(* IEC 61131-3 sources: plc-process-lib/src/POUs/Time/FB_FakeTime, 4 files *)

(* ---- FB_FakeTime.decl.st ---- *)
// Назначение: подменяемый источник времени для тестов: время меняется только вызовами
//             SetNow, Advance, AdvanceL, поэтому тесты таймингов детерминированы и не ждут
//             реального времени. Лежит в библиотеке (не в tests/): им пользуются тесты
//             проектов-потребителей. Старт — LTIME#1H, а не 0: ловит код, который считает
//             «0 = не инициализировано».
// Автор:      kr0nsch
// Версия:     0.1.0
// Документ:   docs/fb/FB_FakeTime.md
FUNCTION_BLOCK FB_FakeTime IMPLEMENTS I_TimeSource
VAR
    ltNow : LTIME := LTIME#1H;   // текущее подменное время
END_VAR

(* ---- Advance.method.decl.st ---- *)
// Продвинуть время на шаг TIME (мс)
METHOD PUBLIC Advance
VAR_INPUT
    tStep : TIME;   // шаг
END_VAR

(* ---- AdvanceL.method.decl.st ---- *)
// Продвинуть время на шаг LTIME: шаги меньше 1 мс и больше 49 сут
METHOD PUBLIC AdvanceL
VAR_INPUT
    ltStep : LTIME;   // шаг
END_VAR

(* ---- SetNow.method.decl.st ---- *)
// Установить время. Можно и назад: ФБ библиотеки обязаны это переживать
METHOD PUBLIC SetNow
VAR_INPUT
    ltValue : LTIME;   // новое время
END_VAR
